Fanuc KAREL source: kt00504.KL

-- PROVISIONAL review KL for V1013-1; original PC SHA256 e17dbafda0a8d3a7c3bedc867876a8db3ba5a4225eb470d8eb06957374713165
-- Incomplete behavior may be omitted. Consult companion uncertainty JSON. Do not deploy.
PROGRAM KT00504
%NOLOCKGROUP
-- UNRESOLVED_DECL P1 type=000102
-- UNRESOLVED_DECL P2 type=000106
-- UNRESOLVED_DECL OUT type=000101
BEGIN
  -- UNRESOLVED_PC offsets 5-20; opcodes 2E,22,32,35
  -- UNRESOLVED_PC offsets 25-40; opcodes 2E,22,32,35
  -- UNRESOLVED_PC offsets 45-79; opcodes 49,7E,49,7E,60,4A
  -- UNRESOLVED_PC offsets 84-88; opcodes 7F
END KT00504
